Fanuc KAREL source: KT00530.KL

PROGRAM KT00530
%NOLOCKGROUP
VAR
  P1: XYZWPREXT
  P2: JOINTPOS
  OUT: XYZWPR
BEGIN
  P1.X = 1.0
  OUT = P1 : P2
END KT00530
